FUNCTION_BLOCK EL_Piston (* The logic of an equipment block: one holder at a time, outputs switched off before new ones go on, all off on release or abort, inputs reported when they change. Technical: Piston: output values from its holder -> outputs (break before make); one holder at a time; all off on release or when the module aborts; inputs -> state channel when they change *)
  (* Standard: 61499-2 *)
  (* Version 0.1, 2026-09-28, Project contributors, AAU Smart Production Lab *)
  PACKAGE stoppering;
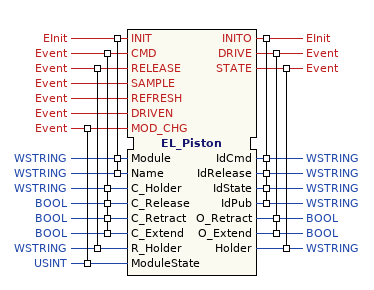
  EVENT_INPUT
    INIT : EInit WITH Module, Name; (* Initialise, once at start-up (the INIT chain); takes the values given with it *)
    CMD WITH C_Holder, C_Release, C_Retract, C_Extend; (* A command arrived from a holder *)
    RELEASE WITH R_Holder; (* A release arrived on the module's release channel (R_Holder) *)
    SAMPLE; (* The inputs were read *)
    REFRESH; (* Cycle: write the outputs again *)
    DRIVEN; (* The outputs were written *)
    MOD_CHG WITH ModuleState; (* The module's state changed (its Aborting switches all off) *)
  END_EVENT
  EVENT_OUTPUT
    INITO : EInit WITH IdCmd, IdRelease, IdState, IdPub; (* Initialised: the next block of the INIT chain goes on *)
    DRIVE WITH O_Retract, O_Extend; (* Write the outputs *)
    STATE WITH Holder; (* Publish the state (the inputs and the holder) *)
  END_EVENT
  VAR_INPUT
    Module : WSTRING; (* The module's name; its local channels are named after it (loc[<Module>/...]) *)
    Name : WSTRING; (* The equipment item's name: its local channels and OPC UA folder *)
    C_Holder : WSTRING; (* Who sends the command *)
    C_Release : BOOL; (* Give up the equipment after this command *)
    C_Retract : BOOL; (* Commanded value of Retract *)
    C_Extend : BOOL; (* Commanded value of Extend *)
    R_Holder : WSTRING; (* Who gives up the equipment *)
    ModuleState : USINT; (* PackML state: 1 Clearing, 2 Stopped, 3 Starting, 4 Idle, 6 Execute, 7 Stopping, 8 Aborting, 9 Aborted, 15 Resetting *)
  END_VAR
  VAR_OUTPUT
    IdCmd : WSTRING; (* Local channel of the commands *)
    IdRelease : WSTRING; (* Local channel of the releases (the module's, one for all equipment) *)
    IdState : WSTRING; (* Local channel of the state *)
    IdPub : WSTRING; (* OPC UA ID of the published inputs *)
    O_Retract : BOOL; (* The value to write to Retract *)
    O_Extend : BOOL; (* The value to write to Extend *)
    Holder : WSTRING; (* Who holds the equipment (empty: free) *)
  END_VAR
  VAR
    Publish : BOOL;
    Beat : USINT;
    LastHolder : WSTRING;
    Pending : BOOL;
    OffPending : BOOL;
    N_Retract : BOOL;
    N_Extend : BOOL;
  END_VAR
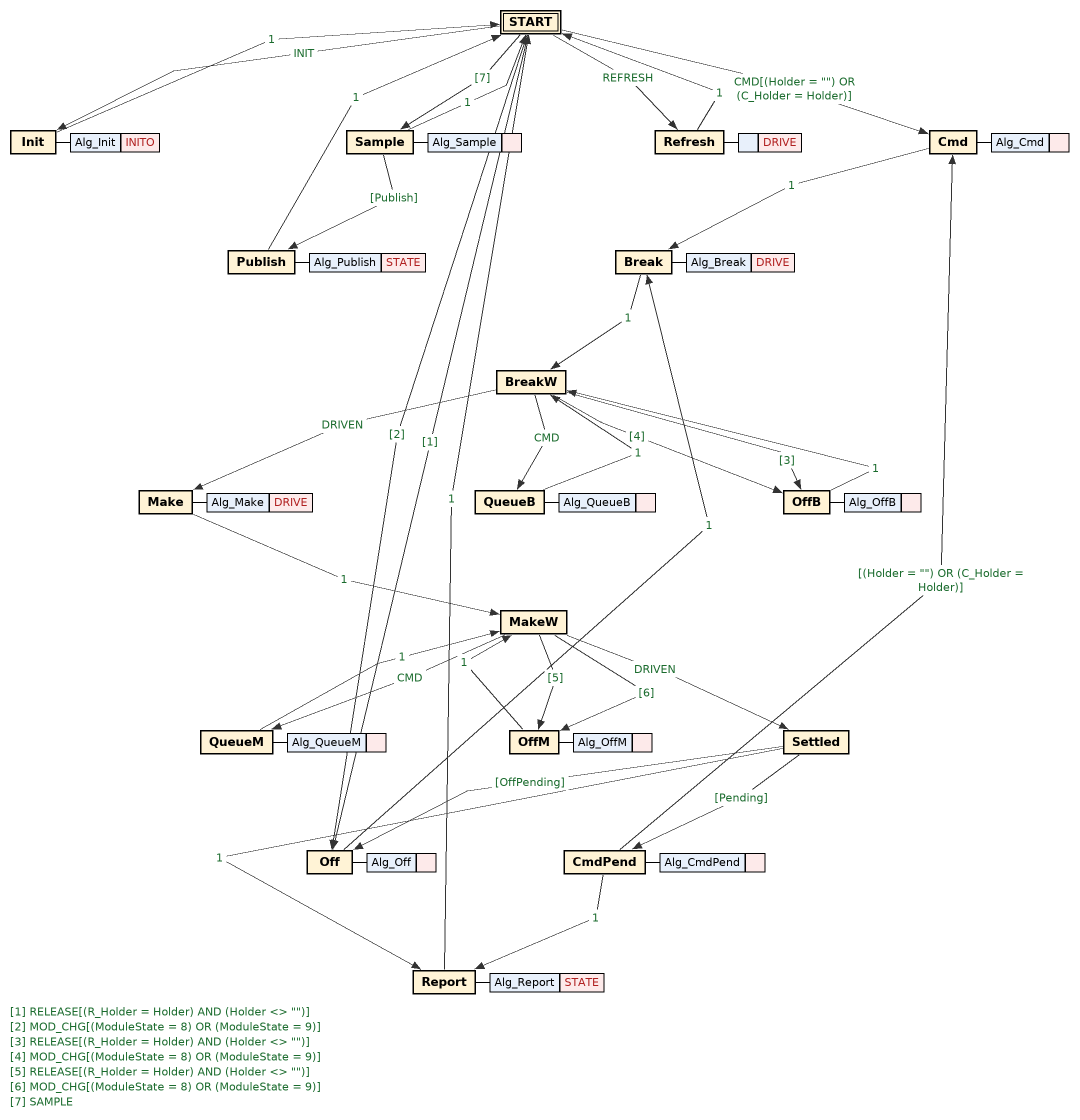
  EC_STATES
    START;
    Init : Alg_Init -> INITO;
    Sample : Alg_Sample;
    Publish : Alg_Publish -> STATE;
    Refresh : -> DRIVE;
    Cmd : Alg_Cmd;
    Off : Alg_Off;
    Break : Alg_Break -> DRIVE;
    Make : Alg_Make -> DRIVE;
    BreakW;
    MakeW;
    QueueB : Alg_QueueB;
    OffB : Alg_OffB;
    QueueM : Alg_QueueM;
    OffM : Alg_OffM;
    CmdPend : Alg_CmdPend;
    Settled;
    Report : Alg_Report -> STATE;
  END_STATES
  EC_TRANSITIONS
    START TO Init := INIT;
    START TO Sample := SAMPLE;
    START TO Refresh := REFRESH;
    START TO Cmd := CMD[(Holder = "") OR (C_Holder = Holder)];
    START TO Off := RELEASE[(R_Holder = Holder) AND (Holder <> "")];
    START TO Off := MOD_CHG[(ModuleState = 8) OR (ModuleState = 9)];
    Init TO START := 1;
    Sample TO Publish := [Publish];
    Sample TO START := 1;
    Publish TO START := 1;
    Refresh TO START := 1;
    Cmd TO Break := 1;
    Off TO Break := 1;
    Break TO BreakW := 1;
    BreakW TO Make := DRIVEN;
    Make TO MakeW := 1;
    MakeW TO Settled := DRIVEN;
    BreakW TO QueueB := CMD;
    BreakW TO OffB := RELEASE[(R_Holder = Holder) AND (Holder <> "")];
    BreakW TO OffB := MOD_CHG[(ModuleState = 8) OR (ModuleState = 9)];
    QueueB TO BreakW := 1;
    OffB TO BreakW := 1;
    MakeW TO QueueM := CMD;
    MakeW TO OffM := RELEASE[(R_Holder = Holder) AND (Holder <> "")];
    MakeW TO OffM := MOD_CHG[(ModuleState = 8) OR (ModuleState = 9)];
    QueueM TO MakeW := 1;
    OffM TO MakeW := 1;
    Settled TO Off := [OffPending];
    Settled TO CmdPend := [Pending];
    CmdPend TO Cmd := [(Holder = "") OR (C_Holder = Holder)];
    CmdPend TO Report := 1;
    Settled TO Report := 1;
    Report TO START := 1;
  END_TRANSITIONS
  ALGORITHM Alg_Init IN ST:
IdCmd := CONCAT(CONCAT(CONCAT(CONCAT("loc[", Module), "/"), Name), "/cmd]");
IdRelease := CONCAT(CONCAT("loc[", Module), "/release]");
IdState := CONCAT(CONCAT(CONCAT(CONCAT("loc[", Module), "/"), Name), "/state]");
IdPub := "";
  END_ALGORITHM
  ALGORITHM Alg_Sample IN ST:
Publish := (Holder <> LastHolder) OR (Beat >= 20);
Beat := Beat + 1;
  END_ALGORITHM
  ALGORITHM Alg_Publish IN ST:
LastHolder := Holder;
Beat := 0;
  END_ALGORITHM
  ALGORITHM Alg_Cmd IN ST:
Holder := C_Holder;
N_Retract := C_Retract;
N_Extend := C_Extend;
IF C_Release THEN
  Holder := "";
END_IF;
  END_ALGORITHM
  ALGORITHM Alg_Off IN ST:
N_Retract := FALSE;
N_Extend := FALSE;
Holder := "";
OffPending := FALSE;
  END_ALGORITHM
  ALGORITHM Alg_Break IN ST:
O_Retract := O_Retract AND N_Retract;
O_Extend := O_Extend AND N_Extend;
  END_ALGORITHM
  ALGORITHM Alg_Make IN ST:
O_Retract := N_Retract;
O_Extend := N_Extend;
  END_ALGORITHM
  ALGORITHM Alg_QueueB IN ST:
Pending := TRUE;
  END_ALGORITHM
  ALGORITHM Alg_OffB IN ST:
OffPending := TRUE;
  END_ALGORITHM
  ALGORITHM Alg_QueueM IN ST:
Pending := TRUE;
  END_ALGORITHM
  ALGORITHM Alg_OffM IN ST:
OffPending := TRUE;
  END_ALGORITHM
  ALGORITHM Alg_CmdPend IN ST:
Pending := FALSE;
  END_ALGORITHM
  ALGORITHM Alg_Report IN ST:
LastHolder := Holder;
Beat := 0;
  END_ALGORITHM
END_FUNCTION_BLOCK
